(* IEC 61131-3 sources: llm-plc-st-eval/data/processed_definitivo/claude-sonnet-4-6/B3/zero_shot, 3 files *)

(* ---- ejec_1.st ---- *)
FUNCTION_BLOCK FB_Contador
VAR_INPUT
    sensorPieza : BOOL; (* Señal del sensor fotoeléctrico *)
    btnReset    : BOOL; (* Botón de reset de cuenta y lote *)
END_VAR

VAR_OUTPUT
    loteListo : BOOL; (* TRUE cuando se alcanzan 12 piezas *)
    cuenta    : INT;  (* Número de piezas contadas *)
END_VAR

VAR
    sensorPiezaAnterior : BOOL; (* Estado previo del sensor para detección de flanco *)
END_VAR

(* ─────────────────────────────────────────────
   Lógica principal
   ───────────────────────────────────────────── *)

(* 1. Reset: tiene prioridad sobre el conteo *)
IF btnReset THEN
    cuenta    := 0;
    loteListo := FALSE;

ELSE
    (* 2. Detección de flanco ascendente del sensor (FALSE → TRUE) *)
    IF sensorPieza AND NOT sensorPiezaAnterior THEN
        cuenta := cuenta + 1;
    END_IF;

    (* 3. Activar salida de lote al alcanzar 12 piezas *)
    IF cuenta >= 12 THEN
        loteListo := TRUE;
    END_IF;

END_IF;

(* 4. Guardar estado actual del sensor para el siguiente ciclo *)
sensorPiezaAnterior := sensorPieza;

(* ---- ejec_2.st ---- *)
FUNCTION_BLOCK FB_Contador
VAR_INPUT
    sensorPieza : BOOL; (* Señal del sensor fotoeléctrico *)
    btnReset    : BOOL; (* Botón de reset de la cuenta *)
END_VAR

VAR_OUTPUT
    loteListo : BOOL; (* Activa cuando se completan 12 piezas *)
    cuenta    : INT;  (* Número de piezas contadas *)
END_VAR

VAR
    sensorPiezaPrev : BOOL; (* Estado anterior del sensor para detección de flanco *)
END_VAR

(*
    Constante de tamaño de lote.
    Ajustar según requerimiento de producción.
*)
VAR CONSTANT
    TAMANO_LOTE : INT := 12;
END_VAR

(* ─────────────────────────────────────────────
   LÓGICA PRINCIPAL
   ───────────────────────────────────────────── *)

(* 1. Reset: tiene prioridad sobre el conteo *)
IF btnReset THEN
    cuenta        := 0;
    loteListo     := FALSE;
    sensorPiezaPrev := FALSE;

ELSE
    (* 2. Detección de flanco ascendente del sensor (FALSE → TRUE) *)
    IF sensorPieza AND NOT sensorPiezaPrev THEN
        (* Incrementar solo si el lote aún no está completo *)
        IF cuenta < TAMANO_LOTE THEN
            cuenta := cuenta + 1;
        END_IF;
    END_IF;

    (* 3. Activar salida de lote completo *)
    IF cuenta >= TAMANO_LOTE THEN
        loteListo := TRUE;
    END_IF;

END_IF;

(* 4. Guardar estado actual del sensor para el siguiente ciclo *)
sensorPiezaPrev := sensorPieza;

END_FUNCTION_BLOCK

(* ---- ejec_3.st ---- *)
FUNCTION_BLOCK FB_Contador
VAR_INPUT
    sensorPieza : BOOL; (* Señal del sensor fotoeléctrico *)
    btnReset    : BOOL; (* Botón de reset de la cuenta *)
END_VAR

VAR_OUTPUT
    loteListo : BOOL; (* Activa cuando se completan 12 piezas *)
    cuenta    : INT;  (* Contador de piezas detectadas *)
END_VAR

VAR
    sensorPiezaPrev : BOOL; (* Estado anterior del sensor para detección de flanco *)
END_VAR

VAR CONSTANT
    LIMITE_LOTE : INT := 12; (* Número de piezas por lote *)
END_VAR

(* ─────────────────────────────────────────────
   Lógica principal del contador de piezas
   ───────────────────────────────────────────── *)

(* 1. Reset: tiene prioridad sobre el conteo *)
IF btnReset THEN
    cuenta    := 0;
    loteListo := FALSE;

(* 2. Conteo: detecta flanco ascendente del sensor (FALSE → TRUE) *)
ELSIF (sensorPieza = TRUE) AND (sensorPiezaPrev = FALSE) THEN

    (* Incrementar solo si el lote aún no está completo *)
    IF cuenta < LIMITE_LOTE THEN
        cuenta := cuenta + 1;
    END_IF;

    (* Activar salida de lote al alcanzar el límite *)
    IF cuenta >= LIMITE_LOTE THEN
        loteListo := TRUE;
    END_IF;

END_IF;

(* 3. Guardar estado actual del sensor para el próximo ciclo *)
sensorPiezaPrev := sensorPieza;
